// TIA Portal V20 export
// export: Created 2026-10-19T18:38:02.6218972Z, ExportSetting WithDefaults, DisplayName Totally Integrated Automation Portal, DisplayVersion V20 Update 6, DisplayName TIA Portal Openness, DisplayVersion V20 Update 6, DisplayName TIA Portal Version Control Interface, DisplayVersion V20 Update 6, DisplayName SINAMICS Startdrive Advanced, DisplayVersion V20 SP1, DisplayName SINAMICS Startdrive G130, G150, S120, S150, SINAMICS MV, G220, S200, S210, DisplayVersion V20 SP1, DisplayName SINAMICS Startdrive G110M, G120, G120C, G120D, G120P, G115D, DisplayVersion V20 SP1, DisplayName STEP 7 Professional, DisplayVersion V20 Update 6, DisplayName STEP 7 Safety, DisplayVersion V20 Update 2, DisplayName WinCC Basic/Comfort/Advanced, DisplayVersion V20 Update 6, DisplayName WinCC Unified, DisplayVersion V20 Update 6
DATA_BLOCK "Order_Table_VTD_FB_DB_1"   // DB6
VERSION : 0.1
// stored: AutoNumber true, DBAccessibleFromOPCUA true, InstanceOfName Order_Table_VTD_FB, InstanceOfType FB
"Order_Table_VTD_FB"
   // VAR_INPUT
   //    System_Selected { ExternalWritable := 'False'} : Bool;
   //    AutoMan_Switch : Bool;
   //    CurrentTime { ExternalWritable := 'False'} : String;
   //    CurrentDTL : DTL;
   //    Watchdog : "Watchdog_Settings_UDT";
   //    VTD_CurrentLevel : UInt;
   //    OPC_UA_State_VTD : UInt;
   //    OPC_UA_state_L2 : UInt;
   //    OPC_UA_state_L3 : UInt;
   //    OPC_UA_state_L4 : UInt;
   //    OPC_UA_state_L5 : UInt;
   //    OPC_UA_state_L6 : UInt;
   //    Clear_OrderTable : Bool;
   // END_VAR
   // VAR_IN_OUT
   //    VTD : "VTD_Control";
   //    Extrator_Conveyor : "ECnv_Control";
   //    Cnv_Buffer_21 : "Buffer_Cnv_Control";
   //    Cnv_Buffer_31 : "Buffer_Cnv_Control";
   //    Cnv_Buffer_41 : "Buffer_Cnv_Control";
   //    Cnv_Buffer_51 : "Buffer_Cnv_Control";
   //    Cnv_Buffer_61 : "Buffer_Cnv_Control";
   //    System : "System_UDT";
   //    Control_OPC_Ua : "WMS_OPC_UA";
   // END_VAR
   // VAR
   //    VTD_CurrentOrder { ExternalWritable := 'False'} : UDInt;
   //    Pallet_InOut_CurrentOrder : UDInt;
   //    Shuttle_InOut_CurrentOrder : UDInt;
   //    VTDDoneRTrig : R_TRIG;
   //    Pallet_InOut_RTrig { S7_SetPoint := 'True'} : R_TRIG;
   //    Shuttle_InOut_RTrig { S7_SetPoint := 'True'} : R_TRIG;
   //    PalletRefused_RTrig { ExternalWritable := 'False'} : R_TRIG;
   //    ErrorRTrig { ExternalWritable := 'False'} : R_TRIG;
   //    CancelRTrig { ExternalWritable := 'False'} : R_TRIG;
   //    PauseRTrig { ExternalWritable := 'False'} : R_TRIG;
   //    ResumeRTrig { ExternalWritable := 'False'} : R_TRIG;
   //    Clear_Store : R_TRIG;
   //    Clear_Retrieve : R_TRIG;
   //    Canceling : Bool;
   //    VTD_WatchdogTimer : TON_TIME;
   //    Pallet_InOut_WatchdogTimer { S7_SetPoint := 'True'} : TON_TIME;
   //    Shuttle_InOut_WatchdogTimer { S7_SetPoint := 'True'} : TON_TIME;
   //    VTD_WatchdogStart : Bool;
   //    Pallet_InOut_WatchdogStart : Bool;
   //    Shuttle_InOut_WatchdogStart : Bool;
   //    F_AutoMode { S7_SetPoint := 'True'} : F_TRIG;
   // END_VAR
BEGIN
END_DATA_BLOCK
